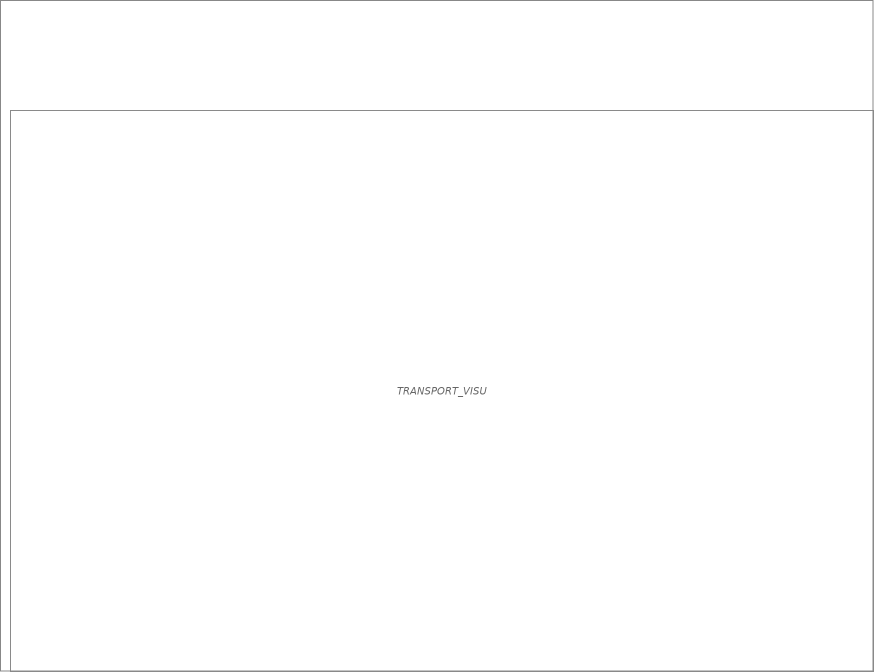
VISUALIZATION MAIN_APPLICATION  // 874x672
    Frame (10,110 864x562)
        shows TRANSPORT_VISU(Data := GVL_APPLICATION.VisuPoolData)
END_VISUALIZATION

(* stored: Version 1.1.0.1, ProductVersion 3.1.4026.20
   Visu MAIN_APPLICATION: Id {c937a261-89d7-4efa-a64e-8edceada3cc4} *)
